Fanuc KAREL source: ka00010.KL

-- PROVISIONAL review KL for V940-1; original PC SHA256 d8515746ab245d5b2e33a169ea169343382885a758eab6548e7ea1cad76dd430
-- Incomplete behavior may be omitted. Consult companion uncertainty JSON. Do not deploy.
PROGRAM KA00010
%NOLOCKGROUP
VAR
  SRC : INTEGER
-- UNRESOLVED_DECL DST type=00001c
BEGIN
  -- V9_ZERO_TABLE_METADATA_HINT layout=0001; no indexed target words; source/name/runtime held
  -- UNRESOLVED_PC offsets 5-16; opcodes 2E,23
  -- UNRESOLVED_PC offsets 21-33; opcodes 21,23
  -- UNRESOLVED_PC offsets 38-42; opcodes 7F
END KA00010
